Fanuc KAREL source: KA00032.KL

PROGRAM KA00032
%NOLOCKGROUP
VAR
  SRC: BOOLEAN
  DST: JOINTPOS
BEGIN
  SRC = TRUE
  DST = SRC
END KA00032
